Yaskawa INFORM job: 11.JBI

/JOB
//NAME 11
//POS
///NPOS 6,6,6,0,0,0
///TOOL 0
///POSTYPE PULSE
///PULSE
C00000=-288,-101153,-84206,3590,-80196,-1936
C00001=6934,-100667,-84028,4379,-80414,-4408
C00002=91626,67370,42890,9351,-80281,-33582
C00003=97267,52739,-6802,12719,-17839,-9459
C00004=137130,47819,-12267,47901,-30619,-34301
C00005=124795,56326,497,57077,-77554,-54431
BC00000=570126
BC00001=225733
BC00002=225733
BC00003=927851
BC00004=927851
BC00005=805226
EC00000=795,0
EC00001=795,0
EC00002=795,0
EC00003=1163,0
EC00004=1163,0
EC00005=795,0
//INST
///DATE 2026/02/11 12:32
///ATTR SC,RW
///GROUP1 RB1,BS1
///GROUP2 ST1
NOP
MOVJ C00000 BC00000 VJ=0.78  +MOVJ EC00000 VJ=0.78
MOVJ C00001 BC00001 VJ=0.78  +MOVJ EC00001 VJ=0.78
MOVJ C00002 BC00002 VJ=0.78  +MOVJ EC00002 VJ=0.78
MOVJ C00003 BC00003 VJ=0.78  +MOVJ EC00003 VJ=0.78
MACRO1 MJ#(0) ARGF1
ARCON
MOVL C00004 BC00004 V=4.2  +MOVJ EC00004 VJ=0.78
WVOF
ARCOF
MOVJ C00005 BC00005 VJ=0.78  +MOVJ EC00005 VJ=0.78
END
